TYPE "ST_LineImage"
VERSION : 0.1
   STRUCT
      LineId : String[40];
      Owner : String[80];
      Revision : UDInt;
      Count : Int;
      Records : Array[1..32] of "ST_LineRecord";
   END_STRUCT;

END_TYPE

